(* IEC 61131-3 sources: avi-aoi-management/knowledge/golden-code/iec61131-st, 3 files *)

(* ---- conveyor-poll-unbounded.st ---- *)
(* Hand-authored STRUCTURALLY-UNSAFE linter golden-corpus example (doc 69 C4; advisory-
   linter demo, not vendor-manual-verified). Certification disclaimer + review process: see
   conveyor-poll-unbounded.meta.md and README.md. *)

(* NEGATIVE example: a condition-driven loop whose condition never turns false and whose
   body has no EXIT/RETURN. Structurally unbounded (an endless scan-cycle loop driving an
   output) even though nothing here names any hazard-domain vocabulary at all — the linter
   flags it on control-flow shape, not wording. *)

PROGRAM ConveyorPoll
VAR
    SensorInput : BOOL;
    MotorRun    : BOOL;
END_VAR

WHILE TRUE DO
    MotorRun := SensorInput;
END_WHILE;

END_PROGRAM

(* ---- debounce-ton.st ---- *)
(* SAFETY: AI-assisted golden example. The author reviews, validates and tests it on a
   simulator before any device runs it. Authors PROCESS logic only; never E-stop /
   interlock / SIL safety functions (those stay on the certified controller).
   See knowledge/golden-code/README.md. *)

PROGRAM DebounceInputSignal
VAR
    RawSignal    : BOOL;             (* noisy field input *)
    DebounceTmr  : TON;              (* standard on-delay timer instance *)
    StableSignal : BOOL;             (* debounced, steady result (output) *)
    DebounceTime : TIME := T#20ms;   (* dwell needed to accept a change *)
END_VAR

(* TON keeps Q low until IN has stayed high past PT (DebounceTime);
   this rejects contact chatter on a mechanical input. *)
DebounceTmr(IN := RawSignal, PT := DebounceTime);
StableSignal := DebounceTmr.Q;

END_PROGRAM

(* ---- moving-average.st ---- *)
(* SAFETY: AI-assisted golden example. The author reviews, validates and tests it on a
   simulator before any device runs it. Authors PROCESS logic only; never E-stop /
   interlock / SIL safety functions (those stay on the certified controller).
   See knowledge/golden-code/README.md. *)

PROGRAM MovingAverage
VAR
    Samples    : ARRAY[0..7] OF REAL;   (* ring buffer, window N = 8 *)
    WriteIndex : INT := 0;              (* next slot to overwrite *)
    Idx        : INT;                   (* cursor over the window *)
    Sum        : REAL := 0.0;
    NewSample  : REAL;                  (* latest raw reading (input) *)
    Average    : REAL;                  (* smoothed result (output) *)
END_VAR

(* push the newest reading into the ring buffer, then advance the cursor *)
Samples[WriteIndex] := NewSample;
WriteIndex := WriteIndex + 1;
IF WriteIndex >= 8 THEN
    WriteIndex := 0;
END_IF;

(* accumulate the whole window, then divide by N *)
Sum := 0.0;
FOR Idx := 0 TO 7 DO
    Sum := Sum + Samples[Idx];
END_FOR;
Average := Sum / 8.0;

END_PROGRAM
